TYPE "DT_DIGITAL_INPUTS_ALL"
VERSION : 0.1
   STRUCT
      CTRL_AND_SYNC : "DT_DIGITAL_INPUT_CTRL_AND_SYNC";
      AUX_SUPPLY : "DT_DIGITAL_INPUT_AUX_SUPPLY";
      GEN_CUBICLE : "DT_DIGITAL_INPUT_GEN_CUBICLE";
      GEN : "DT_DIGITAL_INPUT_GEN";
      PROT : "DT_DIGITAL_INPUT_PROT";
      INTAKE : "DT_DIGITAL_INPUT_INTAKE";
      MIV_AND_BYPASS : "DT_DIGITAL_INPUT_MIV_AND_BYPASS";
      HPU_SYS : "DT_DIGITAL_INPUT_HPU_SYS";
      HPU_PUMPS : "DT_DIGITAL_INPUT_HPU_PUMPS";
      CWS_AND_LOU_SYS : "DT_DIGITAL_INPUT_CWS_AND_LOU_SYS";
      CWS_AND_LOU_PUMPS : "DT_DIGITAL_INPUT_CWS_AND_LOU_PUMPS";
      TURBINE : "DT_DIGITAL_INPUT_TURBINE";
      TRAFO : "DT_DIGITAL_INPUT_TRAFO";
      DRAIN_AND_DEW : "DT_DIGITAL_INPUT_DRAIN_AND_DEW";
      EXC : "DT_DIGITAL_INPUT_EXC";
      SN_LINE : "DT_DIGITAL_INPUT_SN_LINE";
      SN_GEN_AND_MEAS : "DT_DIGITAL_INPUT_SN_GEN_AND_MEAS";
      SN_AUX : "DT_DIGITAL_INPUT_SN_AUX";
      SPARE : "DT_DIGITAL_INPUT_SN_TRAFO";
   END_STRUCT;

END_TYPE

